(* IEC 61131-3 sources: rusty/tests/lit/correctness/control/for, 20 files *)

(* ---- for_loop_evaluates_end_and_step_once_per_iteration.st ---- *)
// RUN: %COMPILE %s && %RUN | %CHECK %s

VAR_GLOBAL
    endCalls, stepCalls : DINT;
END_VAR

FUNCTION getEnd : DINT
    endCalls := endCalls + 1;
    getEnd := 3;
END_FUNCTION

FUNCTION getStep : DINT
    stepCalls := stepCalls + 1;
    getStep := 1;
END_FUNCTION

FUNCTION main : DINT
    VAR
        i, iterations : DINT;
    END_VAR

    // The end and step expressions are evaluated once per iteration and once more to end the loop
    FOR i := 0 TO getEnd() BY getStep() DO
        iterations := iterations + 1;
    END_FOR
    // CHECK: 4 5 5
    printf('%d %d %d$N', iterations, endCalls, stepCalls);
END_FUNCTION

(* ---- continue_in_for_loop_in_while_loop.st ---- *)
// RUN: %COMPILE %s && %RUN | %CHECK %s

FUNCTION main : DINT
    VAR
        i : INT;
    END_VAR

    main := 0;
    WHILE main < 20 DO
        main := main + 1;
        FOR i := 0 TO 10 BY 1 DO
            CONTINUE;
            main := 200;
        END_FOR
    END_WHILE
    main := i + main;

    printf('main=%d$N', main); // CHECK: main=31
END_FUNCTION

(* ---- exit_in_for_loop_in_while_loop.st ---- *)
// RUN: %COMPILE %s && %RUN | %CHECK %s

FUNCTION main : DINT
    VAR
        i : INT;
    END_VAR

    main := 0;
    WHILE main < 20 DO
        main := main + 1;
        FOR i := 0 TO 10 BY 1 DO
            EXIT;
        END_FOR
    END_WHILE
    main := i + main;

    printf('main=%d$N', main); // CHECK: main=20
END_FUNCTION

(* ---- for_continue_test.st ---- *)
// RUN: %COMPILE %s && %RUN | %CHECK %s

FUNCTION main : DINT
    FOR main := 1 TO 10 BY 1 DO
        main := 10;
        CONTINUE;
        main := 200;
    END_FOR

    printf('main=%d$N', main); // CHECK: main=11
END_FUNCTION

(* ---- for_loop_and_decrement_10_times.st ---- *)
// RUN: %COMPILE %s && %RUN | %CHECK %s

FUNCTION main : DINT
    VAR
        i : INT;
    END_VAR

    main := 100;
    FOR i := 10 TO 1 BY -1 DO
        main := main + 1;
    END_FOR

    printf('main=%d$N', main); // CHECK: main=110
END_FUNCTION

(* ---- for_loop_and_increment_10_times.st ---- *)
// RUN: %COMPILE %s && %RUN | %CHECK %s

FUNCTION main : DINT
    VAR
        i : INT;
    END_VAR

    main := 100;
    FOR i := 1 TO 10 DO
        main := main + 1;
    END_FOR

    printf('main=%d$N', main); // CHECK: main=110
END_FUNCTION

(* ---- for_loop_and_increment_10_times_change_vars.st ---- *)
// RUN: %COMPILE %s && %RUN | %CHECK %s

FUNCTION main : DINT
    VAR
        i : INT := 0;
    END_VAR
    VAR_TEMP
        start, end : INT;
    END_VAR

    main := 100;
    start := 1;
    end := 2;
    FOR i := start TO end BY 1 DO
        main := main + 1;
        end := 10;
    END_FOR

    printf('main=%d$N', main); // CHECK: main=110
END_FUNCTION

(* ---- for_loop_and_increment_10_times_skipping_1.st ---- *)
// RUN: %COMPILE %s && %RUN | %CHECK %s

FUNCTION main : DINT
    VAR
        i : INT;
    END_VAR

    main := 1000;
    FOR i := 1 TO 10 BY 2 DO
        main := main + 1;
    END_FOR

    printf('main=%d$N', main); // CHECK: main=1005
END_FUNCTION

(* ---- for_loop_does_not_execute_if_condition_is_not_met.st ---- *)
// RUN: %COMPILE %s && %RUN | %CHECK %s

FUNCTION main : DINT
    VAR
        i, end, step, res : DINT;
    END_VAR

    end := -1;
    step := -1;
    res := 100;

    FOR i := end TO 0 BY step DO
        res := i;
    END_FOR

    main := res;
    printf('main=%d$N', main); // CHECK: main=100
END_FUNCTION

(* ---- for_loop_exit_test.st ---- *)
// RUN: %COMPILE %s && %RUN | %CHECK %s

FUNCTION main : DINT
    FOR main := 100 TO 1000 BY 7 DO
        EXIT;
        main := 200;
    END_FOR

    printf('main=%d$N', main); // CHECK: main=100
END_FUNCTION

(* ---- for_loop_statement_with_binary_expressions.st ---- *)
// RUN: %COMPILE %s && %RUN | %CHECK %s

FUNCTION main : DINT
    VAR
        step : DINT := 1;
        x, y, iteration : DINT;
        z : DINT := 25;
    END_VAR

    // 1 TO 23 BY 3
    FOR x := y + 1 TO z - 2 BY step * 3 DO
        // x: 1, 4, 7, 10, 13, 16, 19, 22
        iteration := iteration + 1;
    END_FOR

    main := iteration;
    printf('main=%d$N', main); // CHECK: main=8
END_FUNCTION

(* ---- for_loop_step_and_counter_change_sign_in_loop_body.st ---- *)
// RUN: %COMPILE %s && %RUN | %CHECK %s

FUNCTION main : DINT
    VAR
        i, step, temp, iteration : DINT;
    END_VAR

    step := 1;
    iteration := 0;

    FOR i := 3 TO 10 BY step DO
        step := (step + 1) * -2;

        // i:     3, -1,   5, -9, 17
        // step: -4,  5, -14, 26
        iteration := iteration + 1;
    END_FOR

    main := iteration;
    printf('main=%d$N', main); // CHECK: main=4
END_FUNCTION

(* ---- for_loop_step_changes_sign_in_loop_body.st ---- *)
// RUN: %COMPILE %s && %RUN | %CHECK %s

FUNCTION main : DINT
    VAR
        i, step, temp, iteration : DINT;
    END_VAR

    step := 1;
    iteration := 0;

    FOR i := 5 TO 10 BY step DO
        temp := (step + 1) * -1;
        IF i + temp > 0 THEN
            step := temp;
        ELSE
            step := step + 3;
        END_IF;

        // i:     5, 3,  4, 2,  3, 1, 2,  6, 1, 5, 12
        // step: -2, 1, -2, 1, -2, 1, 4, -5, 4, 7
        iteration := iteration + 1;
    END_FOR

    main := iteration;
    printf('main=%d$N', main); // CHECK: main=10
END_FUNCTION

(* ---- loop_exit_test.st ---- *)
// RUN: %COMPILE %s && %RUN | %CHECK %s

FUNCTION main : DINT
    FOR main := 100 TO 1000 BY 7 DO
        EXIT;
        main := 200;
    END_FOR
    WHILE main > 50 DO
        EXIT;
        main := 200;
    END_WHILE

    printf('main=%d$N', main); // CHECK: main=100
END_FUNCTION

(* ---- nested_for_loop_allocas_are_hoisted.st ---- *)
// RUN: %COMPILE %s && %RUN | %CHECK %s
//
// Regression test for stack growth caused by lowered loop temporaries.
// Nested FOR loops are desugared into nested WHILE TRUE loops with synthetic
// locals, e.g. roughly:
//
//   alloca __ran_once_1: BOOL
//   alloca __is_incrementing_1: BOOL
//   i := 1
//   __is_incrementing_1 := TRUE
//   WHILE TRUE DO
//       ...
//       alloca __ran_once_0: BOOL
//       alloca __is_incrementing_0: BOOL
//       j := 1
//       __is_incrementing_0 := TRUE
//       WHILE TRUE DO
//           ...
//       END_WHILE
//   END_WHILE
//
// If those `alloca` statements are emitted in-place, the inner loop temps are
// allocated once per outer-loop iteration and the stack eventually overflows at
// `-Onone`. Codegen must hoist the actual stack slots to the function entry
// block and only keep the initialization stores in place.

FUNCTION main : DINT
    VAR
        i, j : DINT;
        counter : DINT;
    END_VAR

    counter := 0;

    FOR i := 1 TO 1000000 DO
        FOR j := 1 TO 1 DO
            counter := counter + 1;
        END_FOR
    END_FOR

    printf('counter=%d$N', counter); // CHECK: counter=1000000
    main := 0;
END_FUNCTION

(* ---- for_loop_overflow.st ---- *)
// RUN: %COMPILE %s && %RUN | %CHECK %s

PROGRAM mainProg
VAR
    i : INT;
    ret : DINT;
END_VAR

ret := 100;
FOR i := 1 TO 0 BY -2 DO
    ret := ret + 1;
END_FOR
END_PROGRAM

FUNCTION main : DINT
    mainProg();

    printf('ret=%d$N', mainProg.ret); // CHECK: ret=101
    printf('i=%d$N', mainProg.i); // CHECK-NEXT: i=-1
    main := 0;
END_FUNCTION

(* ---- for_loop_variable_does_not_affect_other_variables_dint.st ---- *)
// RUN: %COMPILE %s && %RUN | %CHECK %s

PROGRAM mainProg
VAR
    a, i, b, ret : DINT;
END_VAR

a := 16#FFFF_FFFF;
b := 16#FFFF_FFFF;
ret := 100;
FOR i := 1 TO 10 DO
    ret := ret + 1;
END_FOR
END_PROGRAM

FUNCTION main : DINT
    mainProg();

    printf('ret=%d$N', mainProg.ret); // CHECK: ret=110
    printf('a=%d$N', mainProg.a); // CHECK-NEXT: a=-1
    printf('b=%d$N', mainProg.b); // CHECK-NEXT: b=-1
    main := 0;
END_FUNCTION

(* ---- for_loop_variable_does_not_affect_other_variables_int.st ---- *)
// RUN: %COMPILE %s && %RUN | %CHECK %s

PROGRAM mainProg
VAR
    a, i, b : INT;
    ret : DINT;
END_VAR

a := 16#FFFF;
b := 16#FFFF;
ret := 100;
FOR i := 1 TO 10 DO
    ret := ret + 1;
END_FOR
END_PROGRAM

FUNCTION main : DINT
    mainProg();

    printf('ret=%d$N', mainProg.ret); // CHECK: ret=110
    printf('a=%d$N', mainProg.a); // CHECK-NEXT: a=-1
    printf('b=%d$N', mainProg.b); // CHECK-NEXT: b=-1
    main := 0;
END_FUNCTION

(* ---- for_loop_variable_does_not_affect_other_variables_lint.st ---- *)
// RUN: %COMPILE %s && %RUN | %CHECK %s

PROGRAM mainProg
VAR
    a, i, b : LINT;
    ret : DINT;
END_VAR

a := 16#FFFF_FFFF_FFFF_FFFF;
b := 16#FFFF_FFFF_FFFF_FFFF;
ret := 100;
FOR i := 1 TO 10 DO
    ret := ret + 1;
END_FOR
END_PROGRAM

FUNCTION main : DINT
    mainProg();

    printf('ret=%d$N', mainProg.ret); // CHECK: ret=110
    printf('a=%d$N', mainProg.a); // CHECK-NEXT: a=-1
    printf('b=%d$N', mainProg.b); // CHECK-NEXT: b=-1
    main := 0;
END_FUNCTION

(* ---- for_loop_variable_does_not_affect_other_variables_sint.st ---- *)
// RUN: %COMPILE %s && %RUN | %CHECK %s

PROGRAM mainProg
VAR
    a, i, b : SINT;
    ret : DINT;
END_VAR

a := 16#FF;
b := 16#FF;
ret := 100;
FOR i := 1 TO 10 DO
    ret := ret + 1;
END_FOR
END_PROGRAM

FUNCTION main : DINT
    mainProg();

    printf('ret=%d$N', mainProg.ret); // CHECK: ret=110
    printf('a=%d$N', mainProg.a); // CHECK-NEXT: a=-1
    printf('b=%d$N', mainProg.b); // CHECK-NEXT: b=-1
    main := 0;
END_FUNCTION
